Fanuc KAREL source: kt00579.KL

-- PROVISIONAL review KL for V1013-1; original PC SHA256 e6fe6aefe8cfc5a84cf9969060cbece8babc5076caa717ed3dbc39612267cdab
-- Incomplete behavior may be omitted. Consult companion uncertainty JSON. Do not deploy.
PROGRAM KT00579
%NOLOCKGROUP
VAR
  I2 : INTEGER
-- UNRESOLVED_DECL V1 type=000013
-- UNRESOLVED_DECL OUT type=000013
BEGIN
  -- UNRESOLVED_PC offsets 5-20; opcodes 2E,22,32,35
  -- UNRESOLVED_PC offsets 25-36; opcodes 2E,23
  -- UNRESOLVED_PC offsets 41-63; opcodes 49,21,89,4A
  -- UNRESOLVED_PC offsets 68-72; opcodes 7F
END KT00579
